// TIA Portal V20 export
// export: Created 2026-11-20T23:16:57.6278692Z, ExportSetting WithDefaults, DisplayName Totally Integrated Automation Portal, DisplayVersion V20 Update 7, DisplayName TIA Portal Openness, DisplayVersion V20 Update 7, DisplayName TIA Portal Version Control Interface, DisplayVersion V20 Update 7, DisplayName TIA Portal Test Suite Advanced, DisplayVersion V20, DisplayName SINAMICS Startdrive Advanced, DisplayVersion V20 SP1 Update 1, DisplayName SINAMICS Startdrive G110M, G120, G120C, G120D, G120P, G115D, DisplayVersion V20 SP1 Update 1, DisplayName SINAMICS Startdrive G130, G150, S120, S150, SINAMICS MV, G220, S200, S210, DisplayVersion V20 SP1 Update 1, DisplayName STEP 7 Professional, DisplayVersion V20 Update 7, DisplayName STEP 7 Safety, DisplayVersion V20 Update 2, DisplayName WinCC Basic/Comfort/Advanced, DisplayVersion V20 Update 7, DisplayName WinCC Unified, DisplayVersion V20 Update 7
FUNCTION_BLOCK "zzBenSclColours"   // FB260, SCL
{ S7_Optimized_Access := 'TRUE' }
VERSION : 0.1
// stored: AutoNumber true, IsIECCheckEnabled false, IsRetainMemResEnabled false, MemoryReserve 100, SetENOAutomatically false, UDAEnableTagReadback false
   VAR_INPUT
      inEnable : Bool;
      inMode : Int;
      inSetpoint : Real;
   END_VAR
   VAR_OUTPUT
      outActive : Bool;
      outCount : DInt;
      outText : String[40];
   END_VAR
   VAR_IN_OUT
      ioTotal : DInt;
      ioVar : Variant;
   END_VAR
   VAR
      instColFb { S7_SetPoint := 'True'} : "zzBenSclColFb";
      instDelay { S7_SetPoint := 'True'} : TON_TIME;
      statWord : Word;
      statByte : Byte;
      statValues : Array[0..9] of Int;
      statReal : Real;
      statTime : Time;
      statDate : Date;
      statTod : Time_Of_Day;
      statChar : Char;
      statWide : WString[20];
      statFlag : Bool;
      statResult : Int;
      statTimer { S7_SetPoint := 'True'} : IEC_TIMER;
      statÄnderung : Int;
      statÜbung : Int;
   END_VAR
   VAR_TEMP
      tmpI : Int;
      tmpSum : DInt;
      tmpBit : Bool;
   END_VAR
   VAR CONSTANT
      LAST : Int := 9;
   END_VAR
BEGIN
   REGION Constants of each form
       // A line comment on a line of its own
       #statFlag := TRUE;
       #statResult := 42;
       #statResult := -8#17;
       #statWord := 16#00FF;
       #statByte := 2#1010_0101;
       #statReal := 3.14;
       #statReal := 1.5E-3;
       #statTime := T#1s_200ms;
       #statDate := D#2026-11-20;
       #statTod := TOD#12:30:00;
       #statChar := 'A';
       #outText := 'a string with // and (* inside';
       #statWide := WSTRING#'wide';
       #tmpSum := DINT#-7;
       #statWord := WORD#16#0F0F;
   END_REGION

   REGION Operands
       (* A block comment
          over two lines *)
       #outActive := #inEnable AND "zzMcTag1"; // a comment after code
       "zzBenSclColDb".motor.speed := #inMode;
       "zzBenSclColDb".values[#tmpI] := #statValues[LAST];
       #tmpBit := #statWord.%X3;
       #statByte := #statWord.%B0;
       #ioTotal += #outCount;
       "zzMcTag1" := #tmpBit;
   END_REGION

   REGION Keywords
       IF #inMode = 1 THEN
           #statResult := 1;
       ELSIF #inMode > 1 AND #inMode <= 5 THEN
           #statResult := #inMode MOD 2;
       ELSE
           #statResult := 0;
       END_IF;

       CASE #inMode OF
           0:
               #outText := 'idle';
           1..3, 5:
               #outText := 'run';
           ELSE
               #outText := '';
       END_CASE;

       #tmpSum := 0;
       FOR #tmpI := 0 TO #LAST BY 1 DO
           IF #statValues[#tmpI] < 0 THEN
               CONTINUE;
           END_IF;
           #tmpSum := #tmpSum + #statValues[#tmpI];
           IF #tmpSum > 1000 THEN
               EXIT;
           END_IF;
       END_FOR;

       #tmpI := 0;
       WHILE #tmpI < #LAST AND NOT #statFlag DO
           #tmpI := #tmpI + 1;
       END_WHILE;

       REPEAT
           #tmpI := #tmpI - 1;
       UNTIL #tmpI <= 0 OR #statFlag XOR #tmpBit
       END_REPEAT;
   END_REGION

   REGION Calls
       // An instruction with an instance and without, an FC, an FB as a multi-instance and with its DB
       #instDelay(IN := #inEnable,
                  PT := T#5s,
                  Q => #statFlag,
                  ET => #statTime);
       #statResult := MAX(IN1 := #statResult, IN2 := 10);
       #statReal := SQRT(ABS(#inSetpoint)) ** 2.0;
       #statResult := "zzBenSclColFc"(inA := #statResult, inB := 5);
       #instColFb(inStart := #statFlag,
                  outDone => #tmpBit);
       "zzBenSclColFbDb"(inStart := #inEnable);
       #outCount := INT_TO_DINT(#statResult) * 2 - #tmpSum / 3;
   END_REGION

   REGION Settled by TIA // a comment on the region's line
       (/*A multilingual comment in code*/)
       ENO := FALSE;
       IF TypeOf(#ioVar) = Int THEN
           #statÄnderung := 1;
       ELSIF TypeOf(#ioVar) = zzBenSclColType THEN
           #statÄnderung := 2;
       END_IF;
       #statTimer.TON(IN := #inEnable, PT := T#2s);
       #statÜbung := #statÄnderung + 1;
   END_REGION

   IF NOT #inEnable THEN
       GOTO lblEnd;
   END_IF;
   #outActive := #instColFb.outDone OR "zzBenSclColFbDb".outDone;
   RETURN;
   lblEnd: #outActive := FALSE;
END_FUNCTION_BLOCK
